# EPICS substitutions: b-55B2VNC/src/main/epics/PCF5CoreApp/Db/Oscil_NDS_StateMachine.substitutions
file "nds3_StateMachine.template"{
pattern
{
    BOARDTYPE,
    BOARDTYPEIDX,
    CBS1,
    CBS2,
    STATEMACHINE_PARENT,
    STATEMACHINE_NAME
}
{
    "B",
    "7",
    "D1",
    "I2",
    "",
    "StateMachine"
}
}
